Fanuc KAREL source: KT00926.KL

PROGRAM KT00926
%NOLOCKGROUP
VAR
  Y1: ARRAY[2] OF BYTE
  Y2: ARRAY[2] OF BYTE
  OUT: STRING[80]
BEGIN
  Y1[1] = 2
  Y2[1] = 3
  Y1[1] = 2
  Y2[1] = 3
  OUT = SUB_STR(Y1[1], 1, 1)
END KT00926
